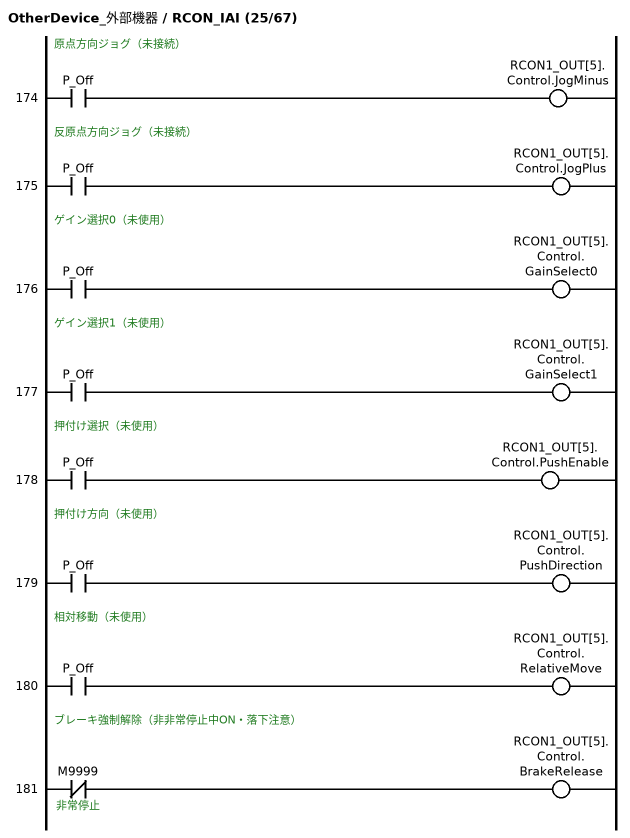
(* [picture p96: OtherDevice_外部機器 / RCON_IAI, rungs 174-181] *)
(* Rung 174: 原点方向ジョグ（未接続） *)
RCON1_OUT[5].Control.JogMinus := P_Off;
(* Rung 175: 反原点方向ジョグ（未接続） *)
RCON1_OUT[5].Control.JogPlus := P_Off;
(* Rung 176: ゲイン選択0（未使用） *)
RCON1_OUT[5].Control.GainSelect0 := P_Off;
(* Rung 177: ゲイン選択1（未使用） *)
RCON1_OUT[5].Control.GainSelect1 := P_Off;
(* Rung 178: 押付け選択（未使用） *)
RCON1_OUT[5].Control.PushEnable := P_Off;
(* Rung 179: 押付け方向（未使用） *)
RCON1_OUT[5].Control.PushDirection := P_Off;
(* Rung 180: 相対移動（未使用） *)
RCON1_OUT[5].Control.RelativeMove := P_Off;
(* Rung 181: ブレーキ強制解除（非非常停止中ON・落下注意） *)
RCON1_OUT[5].Control.BrakeRelease := NOT M9999;

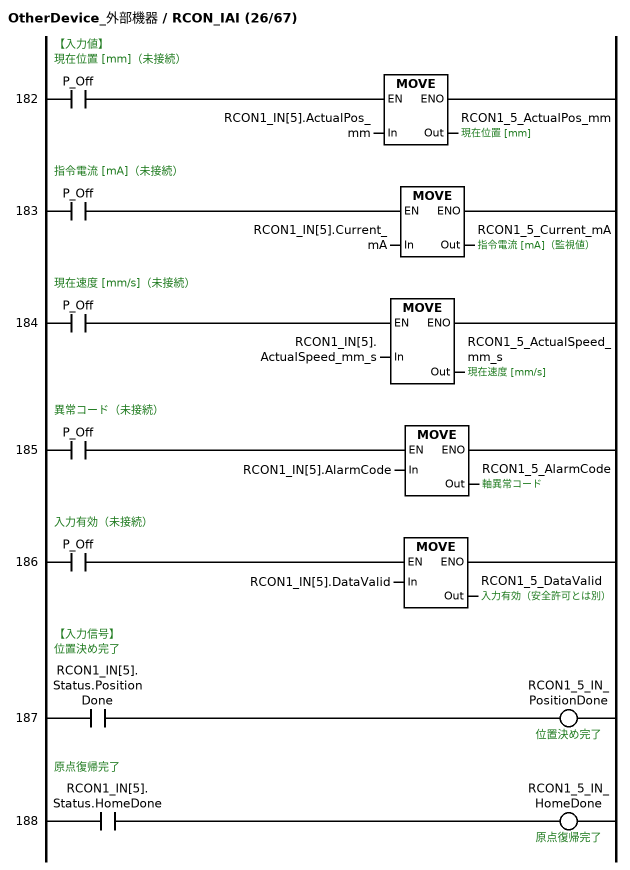
(* Rung 182: 【入力値】 / 現在位置 [mm]（未接続） *)
IF P_Off THEN RCON1_5_ActualPos_mm := RCON1_IN[5].ActualPos_mm; END_IF;
(* Rung 183: 指令電流 [mA]（未接続） *)
IF P_Off THEN RCON1_5_Current_mA := RCON1_IN[5].Current_mA; END_IF;
(* Rung 184: 現在速度 [mm/s]（未接続） *)
IF P_Off THEN RCON1_5_ActualSpeed_mm_s := RCON1_IN[5].ActualSpeed_mm_s; END_IF;
(* Rung 185: 異常コード（未接続） *)
IF P_Off THEN RCON1_5_AlarmCode := RCON1_IN[5].AlarmCode; END_IF;
(* Rung 186: 入力有効（未接続） *)
IF P_Off THEN RCON1_5_DataValid := RCON1_IN[5].DataValid; END_IF;
(* Rung 187: 【入力信号】 / 位置決め完了 *)
RCON1_5_IN_PositionDone := RCON1_IN[5].Status.PositionDone;
(* Rung 188: 原点復帰完了 *)
RCON1_5_IN_HomeDone := RCON1_IN[5].Status.HomeDone;

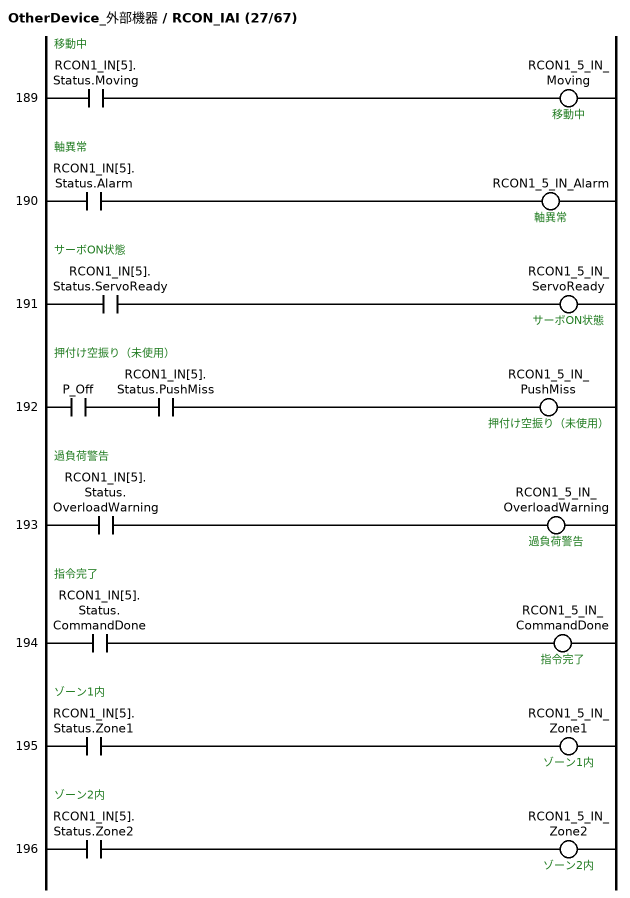
(* Rung 189: 移動中 *)
RCON1_5_IN_Moving := RCON1_IN[5].Status.Moving;
(* Rung 190: 軸異常 *)
RCON1_5_IN_Alarm := RCON1_IN[5].Status.Alarm;
(* Rung 191: サーボON状態 *)
RCON1_5_IN_ServoReady := RCON1_IN[5].Status.ServoReady;
(* Rung 192: 押付け空振り（未使用） *)
RCON1_5_IN_PushMiss := P_Off AND RCON1_IN[5].Status.PushMiss;
(* Rung 193: 過負荷警告 *)
RCON1_5_IN_OverloadWarning := RCON1_IN[5].Status.OverloadWarning;
(* Rung 194: 指令完了 *)
RCON1_5_IN_CommandDone := RCON1_IN[5].Status.CommandDone;
(* Rung 195: ゾーン1内 *)
RCON1_5_IN_Zone1 := RCON1_IN[5].Status.Zone1;
(* Rung 196: ゾーン2内 *)
RCON1_5_IN_Zone2 := RCON1_IN[5].Status.Zone2;

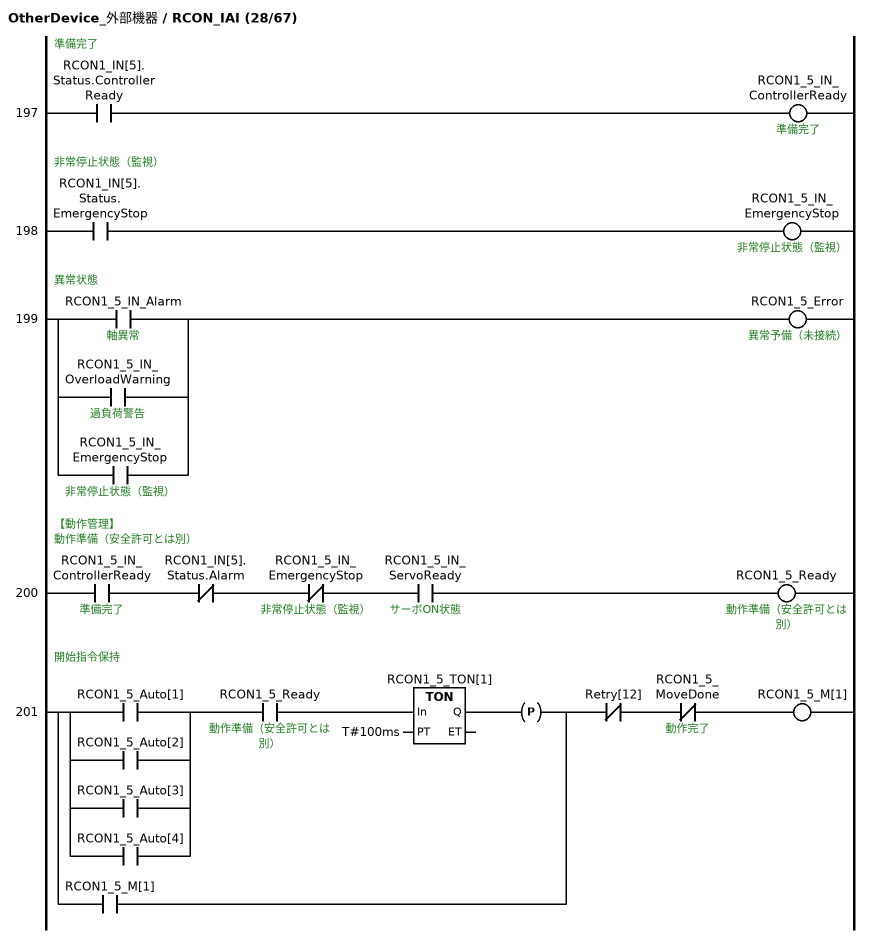
(* Rung 197: 準備完了 *)
RCON1_5_IN_ControllerReady := RCON1_IN[5].Status.ControllerReady;
(* Rung 198: 非常停止状態（監視） *)
RCON1_5_IN_EmergencyStop := RCON1_IN[5].Status.EmergencyStop;
(* Rung 199: 異常状態 *)
RCON1_5_Error := RCON1_5_IN_Alarm OR RCON1_5_IN_OverloadWarning OR RCON1_5_IN_EmergencyStop;
(* Rung 200: 【動作管理】 / 動作準備（安全許可とは別） *)
RCON1_5_Ready := RCON1_5_IN_ControllerReady AND NOT RCON1_IN[5].Status.Alarm AND NOT RCON1_5_IN_EmergencyStop AND RCON1_5_IN_ServoReady;
(* Rung 201: 開始指令保持 *)
RCON1_5_TON[1](In := (RCON1_5_Auto[1] OR RCON1_5_Auto[2] OR RCON1_5_Auto[3] OR RCON1_5_Auto[4]) AND RCON1_5_Ready, PT := T#100ms);
_e18(CLK := RCON1_5_TON[1].Q);
RCON1_5_M[1] := (_e18.Q OR RCON1_5_M[1]) AND NOT Retry[12] AND NOT RCON1_5_MoveDone;

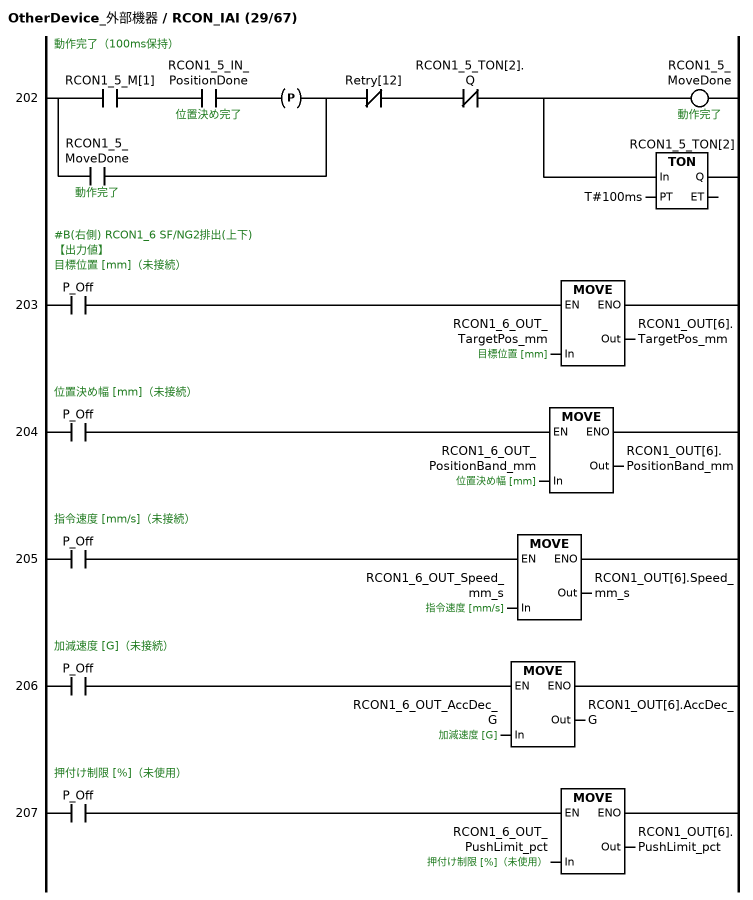
(* Rung 202: 動作完了（100ms保持） *)
_e19(CLK := RCON1_5_M[1] AND RCON1_5_IN_PositionDone);
_p20 := (_e19.Q OR RCON1_5_MoveDone) AND NOT Retry[12] AND NOT RCON1_5_TON[2].Q;
RCON1_5_MoveDone := _p20;
RCON1_5_TON[2](In := _p20, PT := T#100ms);
(* Rung 203: #B(右側) RCON1_6 SF/NG2排出(上下) / 【出力値】 / 目標位置 [mm]（未接続） *)
IF P_Off THEN RCON1_OUT[6].TargetPos_mm := RCON1_6_OUT_TargetPos_mm; END_IF;
(* Rung 204: 位置決め幅 [mm]（未接続） *)
IF P_Off THEN RCON1_OUT[6].PositionBand_mm := RCON1_6_OUT_PositionBand_mm; END_IF;
(* Rung 205: 指令速度 [mm/s]（未接続） *)
IF P_Off THEN RCON1_OUT[6].Speed_mm_s := RCON1_6_OUT_Speed_mm_s; END_IF;
(* Rung 206: 加減速度 [G]（未接続） *)
IF P_Off THEN RCON1_OUT[6].AccDec_G := RCON1_6_OUT_AccDec_G; END_IF;
(* Rung 207: 押付け制限 [%]（未使用） *)
IF P_Off THEN RCON1_OUT[6].PushLimit_pct := RCON1_6_OUT_PushLimit_pct; END_IF;

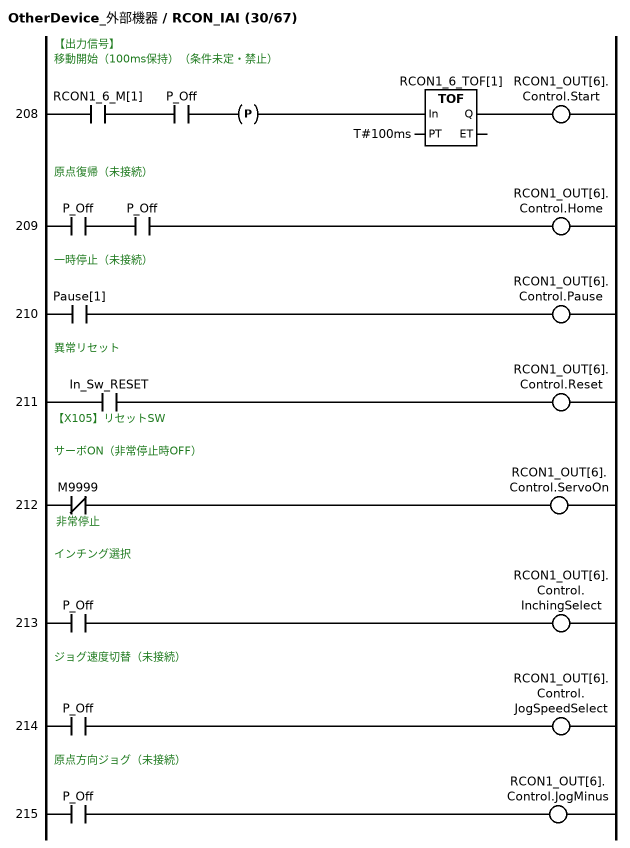
(* Rung 208: 【出力信号】 / 移動開始（100ms保持）（条件未定・禁止） *)
_e21(CLK := RCON1_6_M[1] AND P_Off);
RCON1_6_TOF[1](In := _e21.Q, PT := T#100ms);
RCON1_OUT[6].Control.Start := RCON1_6_TOF[1].Q;
(* Rung 209: 原点復帰（未接続） *)
RCON1_OUT[6].Control.Home := P_Off AND P_Off;
(* Rung 210: 一時停止（未接続） *)
RCON1_OUT[6].Control.Pause := Pause[1];
(* Rung 211: 異常リセット *)
RCON1_OUT[6].Control.Reset := In_Sw_RESET;
(* Rung 212: サーボON（非常停止時OFF） *)
RCON1_OUT[6].Control.ServoOn := NOT M9999;
(* Rung 213: インチング選択 *)
RCON1_OUT[6].Control.InchingSelect := P_Off;
(* Rung 214: ジョグ速度切替（未接続） *)
RCON1_OUT[6].Control.JogSpeedSelect := P_Off;
(* Rung 215: 原点方向ジョグ（未接続） *)
RCON1_OUT[6].Control.JogMinus := P_Off;

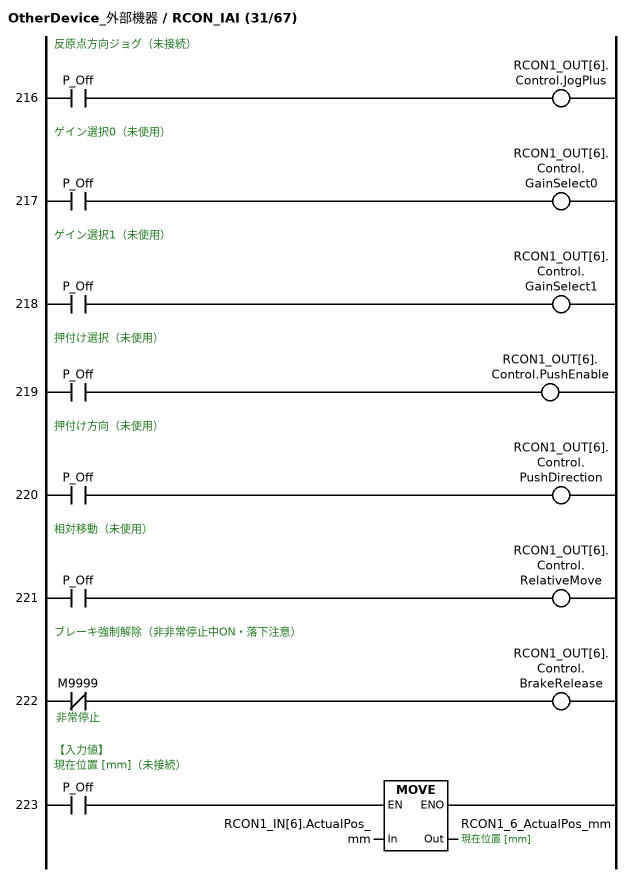
(* Rung 216: 反原点方向ジョグ（未接続） *)
RCON1_OUT[6].Control.JogPlus := P_Off;
(* Rung 217: ゲイン選択0（未使用） *)
RCON1_OUT[6].Control.GainSelect0 := P_Off;
(* Rung 218: ゲイン選択1（未使用） *)
RCON1_OUT[6].Control.GainSelect1 := P_Off;
(* Rung 219: 押付け選択（未使用） *)
RCON1_OUT[6].Control.PushEnable := P_Off;
(* Rung 220: 押付け方向（未使用） *)
RCON1_OUT[6].Control.PushDirection := P_Off;
(* Rung 221: 相対移動（未使用） *)
RCON1_OUT[6].Control.RelativeMove := P_Off;
(* Rung 222: ブレーキ強制解除（非非常停止中ON・落下注意） *)
RCON1_OUT[6].Control.BrakeRelease := NOT M9999;
(* Rung 223: 【入力値】 / 現在位置 [mm]（未接続） *)
IF P_Off THEN RCON1_6_ActualPos_mm := RCON1_IN[6].ActualPos_mm; END_IF;

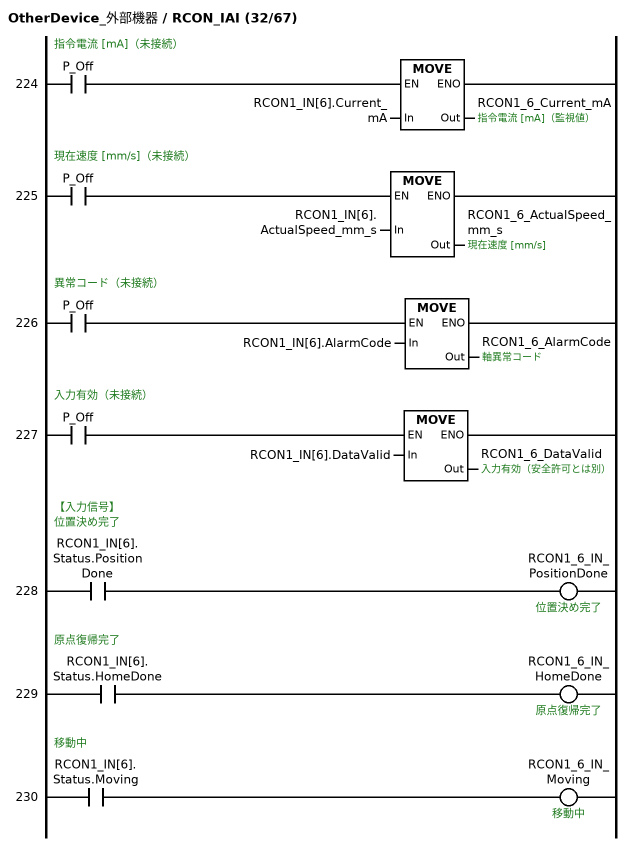
(* Rung 224: 指令電流 [mA]（未接続） *)
IF P_Off THEN RCON1_6_Current_mA := RCON1_IN[6].Current_mA; END_IF;
(* Rung 225: 現在速度 [mm/s]（未接続） *)
IF P_Off THEN RCON1_6_ActualSpeed_mm_s := RCON1_IN[6].ActualSpeed_mm_s; END_IF;
(* Rung 226: 異常コード（未接続） *)
IF P_Off THEN RCON1_6_AlarmCode := RCON1_IN[6].AlarmCode; END_IF;
(* Rung 227: 入力有効（未接続） *)
IF P_Off THEN RCON1_6_DataValid := RCON1_IN[6].DataValid; END_IF;
(* Rung 228: 【入力信号】 / 位置決め完了 *)
RCON1_6_IN_PositionDone := RCON1_IN[6].Status.PositionDone;
(* Rung 229: 原点復帰完了 *)
RCON1_6_IN_HomeDone := RCON1_IN[6].Status.HomeDone;
(* Rung 230: 移動中 *)
RCON1_6_IN_Moving := RCON1_IN[6].Status.Moving;

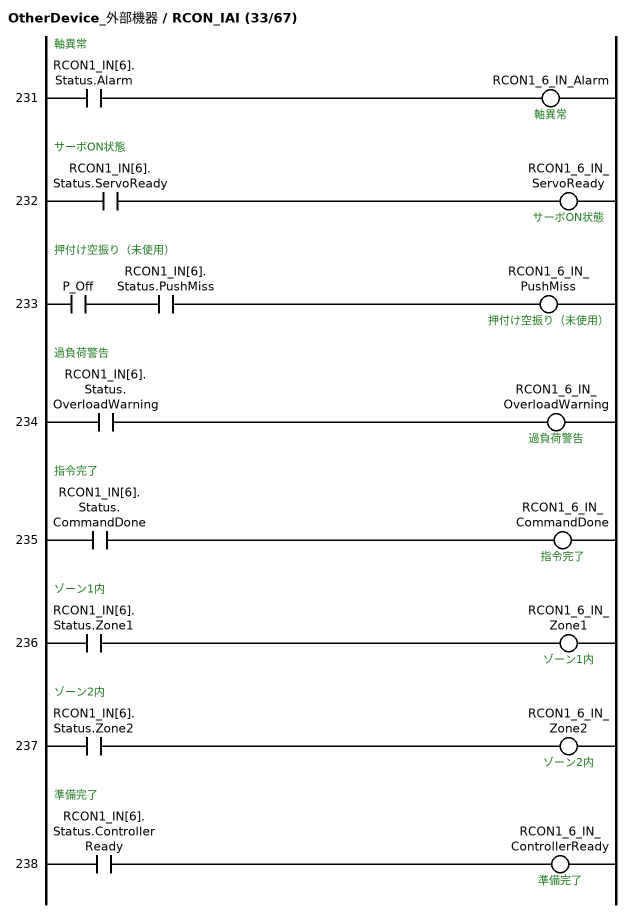
(* Rung 231: 軸異常 *)
RCON1_6_IN_Alarm := RCON1_IN[6].Status.Alarm;
(* Rung 232: サーボON状態 *)
RCON1_6_IN_ServoReady := RCON1_IN[6].Status.ServoReady;
(* Rung 233: 押付け空振り（未使用） *)
RCON1_6_IN_PushMiss := P_Off AND RCON1_IN[6].Status.PushMiss;
(* Rung 234: 過負荷警告 *)
RCON1_6_IN_OverloadWarning := RCON1_IN[6].Status.OverloadWarning;
(* Rung 235: 指令完了 *)
RCON1_6_IN_CommandDone := RCON1_IN[6].Status.CommandDone;
(* Rung 236: ゾーン1内 *)
RCON1_6_IN_Zone1 := RCON1_IN[6].Status.Zone1;
(* Rung 237: ゾーン2内 *)
RCON1_6_IN_Zone2 := RCON1_IN[6].Status.Zone2;
(* Rung 238: 準備完了 *)
RCON1_6_IN_ControllerReady := RCON1_IN[6].Status.ControllerReady;

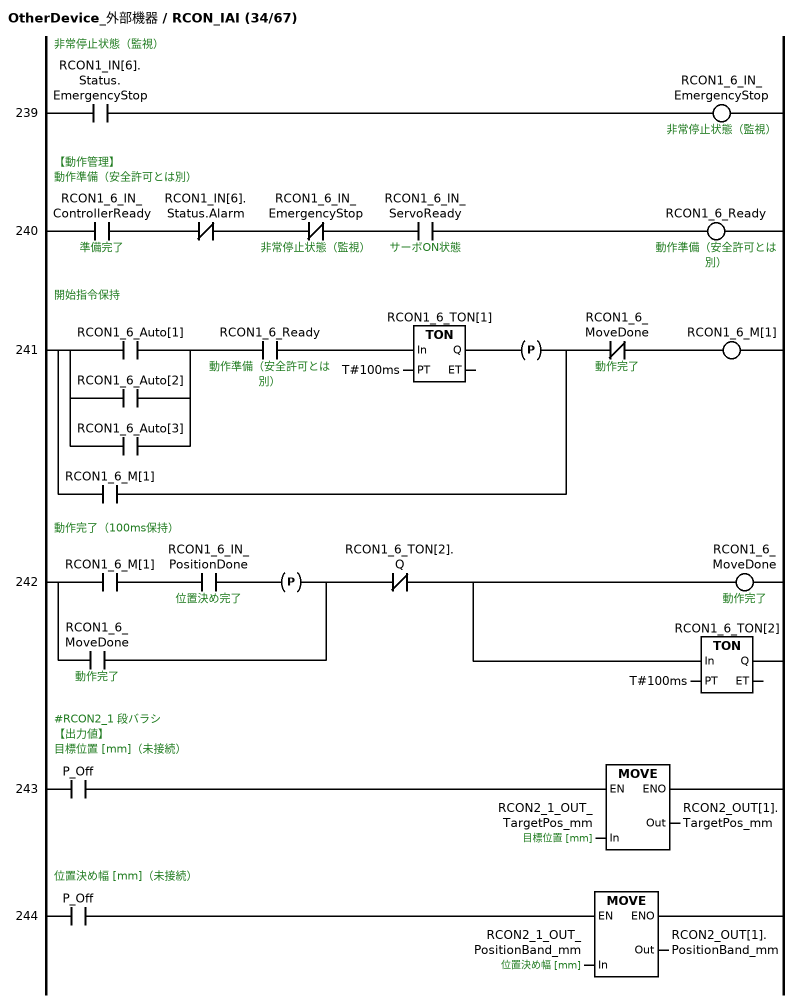
(* Rung 239: 非常停止状態（監視） *)
RCON1_6_IN_EmergencyStop := RCON1_IN[6].Status.EmergencyStop;
(* Rung 240: 【動作管理】 / 動作準備（安全許可とは別） *)
RCON1_6_Ready := RCON1_6_IN_ControllerReady AND NOT RCON1_IN[6].Status.Alarm AND NOT RCON1_6_IN_EmergencyStop AND RCON1_6_IN_ServoReady;
(* Rung 241: 開始指令保持 *)
RCON1_6_TON[1](In := (RCON1_6_Auto[1] OR RCON1_6_Auto[2] OR RCON1_6_Auto[3]) AND RCON1_6_Ready, PT := T#100ms);
_e22(CLK := RCON1_6_TON[1].Q);
RCON1_6_M[1] := (_e22.Q OR RCON1_6_M[1]) AND NOT RCON1_6_MoveDone;
(* Rung 242: 動作完了（100ms保持） *)
_e23(CLK := RCON1_6_M[1] AND RCON1_6_IN_PositionDone);
_p24 := (_e23.Q OR RCON1_6_MoveDone) AND NOT RCON1_6_TON[2].Q;
RCON1_6_MoveDone := _p24;
RCON1_6_TON[2](In := _p24, PT := T#100ms);
(* Rung 243: #RCON2_1 段バラシ / 【出力値】 / 目標位置 [mm]（未接続） *)
IF P_Off THEN RCON2_OUT[1].TargetPos_mm := RCON2_1_OUT_TargetPos_mm; END_IF;
(* Rung 244: 位置決め幅 [mm]（未接続） *)
IF P_Off THEN RCON2_OUT[1].PositionBand_mm := RCON2_1_OUT_PositionBand_mm; END_IF;

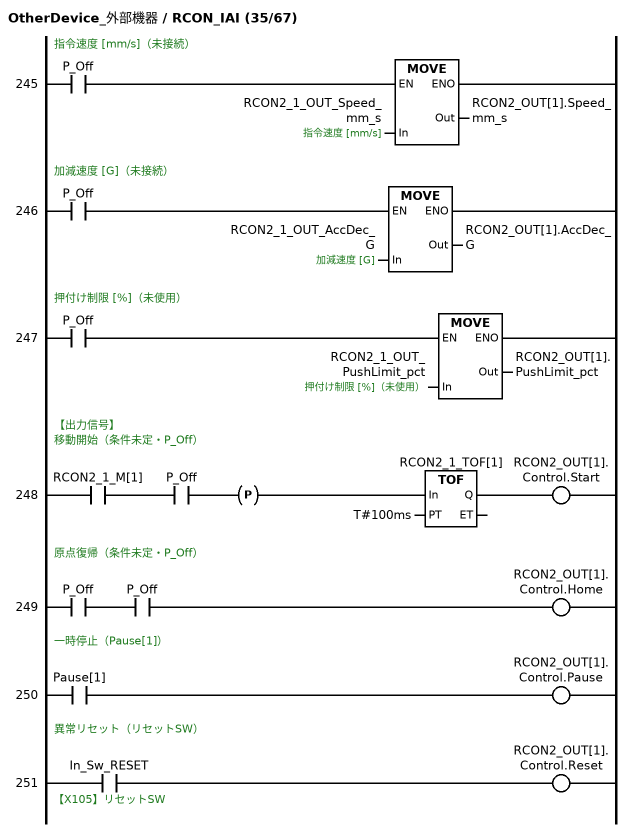
(* Rung 245: 指令速度 [mm/s]（未接続） *)
IF P_Off THEN RCON2_OUT[1].Speed_mm_s := RCON2_1_OUT_Speed_mm_s; END_IF;
(* Rung 246: 加減速度 [G]（未接続） *)
IF P_Off THEN RCON2_OUT[1].AccDec_G := RCON2_1_OUT_AccDec_G; END_IF;
(* Rung 247: 押付け制限 [%]（未使用） *)
IF P_Off THEN RCON2_OUT[1].PushLimit_pct := RCON2_1_OUT_PushLimit_pct; END_IF;
(* Rung 248: 【出力信号】 / 移動開始（条件未定・P_Off） *)
_e25(CLK := RCON2_1_M[1] AND P_Off);
RCON2_1_TOF[1](In := _e25.Q, PT := T#100ms);
RCON2_OUT[1].Control.Start := RCON2_1_TOF[1].Q;
(* Rung 249: 原点復帰（条件未定・P_Off） *)
RCON2_OUT[1].Control.Home := P_Off AND P_Off;
(* Rung 250: 一時停止（Pause[1]） *)
RCON2_OUT[1].Control.Pause := Pause[1];
(* Rung 251: 異常リセット（リセットSW） *)
RCON2_OUT[1].Control.Reset := In_Sw_RESET;

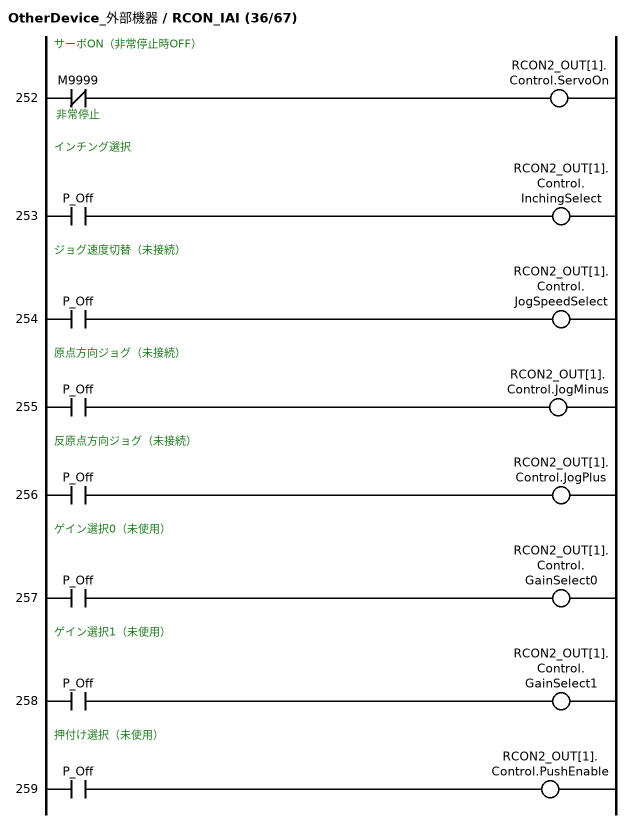
(* Rung 252: サーボON（非常停止時OFF） *)
RCON2_OUT[1].Control.ServoOn := NOT M9999;
(* Rung 253: インチング選択 *)
RCON2_OUT[1].Control.InchingSelect := P_Off;
(* Rung 254: ジョグ速度切替（未接続） *)
RCON2_OUT[1].Control.JogSpeedSelect := P_Off;
(* Rung 255: 原点方向ジョグ（未接続） *)
RCON2_OUT[1].Control.JogMinus := P_Off;
(* Rung 256: 反原点方向ジョグ（未接続） *)
RCON2_OUT[1].Control.JogPlus := P_Off;
(* Rung 257: ゲイン選択0（未使用） *)
RCON2_OUT[1].Control.GainSelect0 := P_Off;
(* Rung 258: ゲイン選択1（未使用） *)
RCON2_OUT[1].Control.GainSelect1 := P_Off;
(* Rung 259: 押付け選択（未使用） *)
RCON2_OUT[1].Control.PushEnable := P_Off;

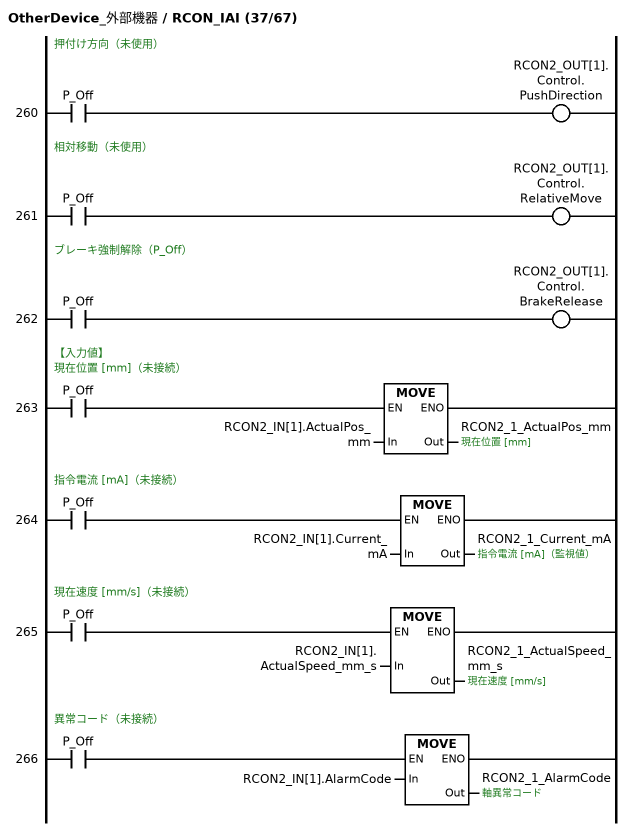
(* Rung 260: 押付け方向（未使用） *)
RCON2_OUT[1].Control.PushDirection := P_Off;
(* Rung 261: 相対移動（未使用） *)
RCON2_OUT[1].Control.RelativeMove := P_Off;
(* Rung 262: ブレーキ強制解除（P_Off） *)
RCON2_OUT[1].Control.BrakeRelease := P_Off;
(* Rung 263: 【入力値】 / 現在位置 [mm]（未接続） *)
IF P_Off THEN RCON2_1_ActualPos_mm := RCON2_IN[1].ActualPos_mm; END_IF;
(* Rung 264: 指令電流 [mA]（未接続） *)
IF P_Off THEN RCON2_1_Current_mA := RCON2_IN[1].Current_mA; END_IF;
(* Rung 265: 現在速度 [mm/s]（未接続） *)
IF P_Off THEN RCON2_1_ActualSpeed_mm_s := RCON2_IN[1].ActualSpeed_mm_s; END_IF;
(* Rung 266: 異常コード（未接続） *)
IF P_Off THEN RCON2_1_AlarmCode := RCON2_IN[1].AlarmCode; END_IF;

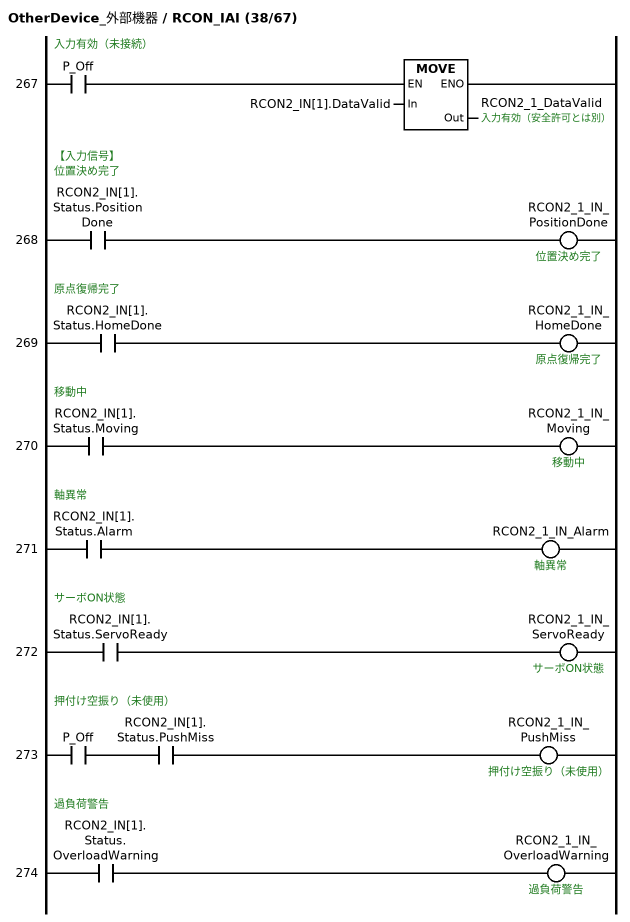
(* Rung 267: 入力有効（未接続） *)
IF P_Off THEN RCON2_1_DataValid := RCON2_IN[1].DataValid; END_IF;
(* Rung 268: 【入力信号】 / 位置決め完了 *)
RCON2_1_IN_PositionDone := RCON2_IN[1].Status.PositionDone;
(* Rung 269: 原点復帰完了 *)
RCON2_1_IN_HomeDone := RCON2_IN[1].Status.HomeDone;
(* Rung 270: 移動中 *)
RCON2_1_IN_Moving := RCON2_IN[1].Status.Moving;
(* Rung 271: 軸異常 *)
RCON2_1_IN_Alarm := RCON2_IN[1].Status.Alarm;
(* Rung 272: サーボON状態 *)
RCON2_1_IN_ServoReady := RCON2_IN[1].Status.ServoReady;
(* Rung 273: 押付け空振り（未使用） *)
RCON2_1_IN_PushMiss := P_Off AND RCON2_IN[1].Status.PushMiss;
(* Rung 274: 過負荷警告 *)
RCON2_1_IN_OverloadWarning := RCON2_IN[1].Status.OverloadWarning;

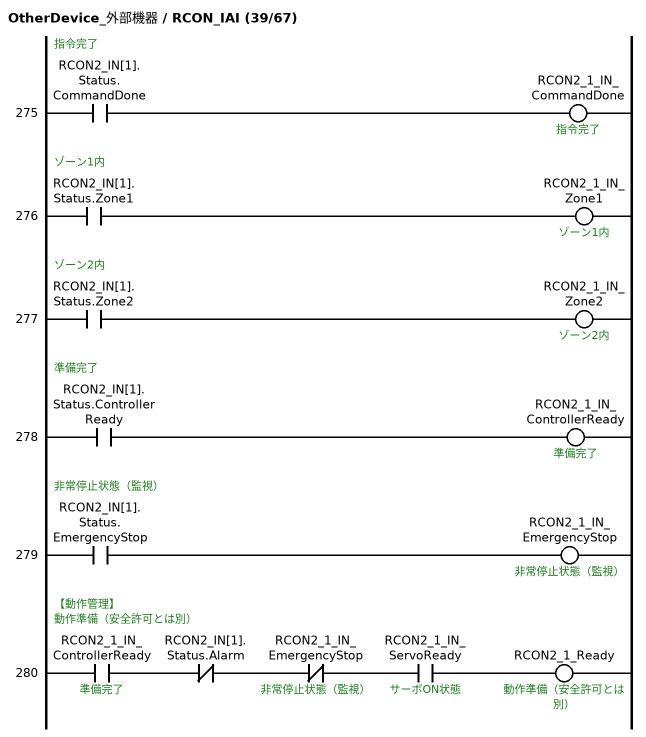
(* Rung 275: 指令完了 *)
RCON2_1_IN_CommandDone := RCON2_IN[1].Status.CommandDone;
(* Rung 276: ゾーン1内 *)
RCON2_1_IN_Zone1 := RCON2_IN[1].Status.Zone1;
(* Rung 277: ゾーン2内 *)
RCON2_1_IN_Zone2 := RCON2_IN[1].Status.Zone2;
(* Rung 278: 準備完了 *)
RCON2_1_IN_ControllerReady := RCON2_IN[1].Status.ControllerReady;
(* Rung 279: 非常停止状態（監視） *)
RCON2_1_IN_EmergencyStop := RCON2_IN[1].Status.EmergencyStop;
(* Rung 280: 【動作管理】 / 動作準備（安全許可とは別） *)
RCON2_1_Ready := RCON2_1_IN_ControllerReady AND NOT RCON2_IN[1].Status.Alarm AND NOT RCON2_1_IN_EmergencyStop AND RCON2_1_IN_ServoReady;

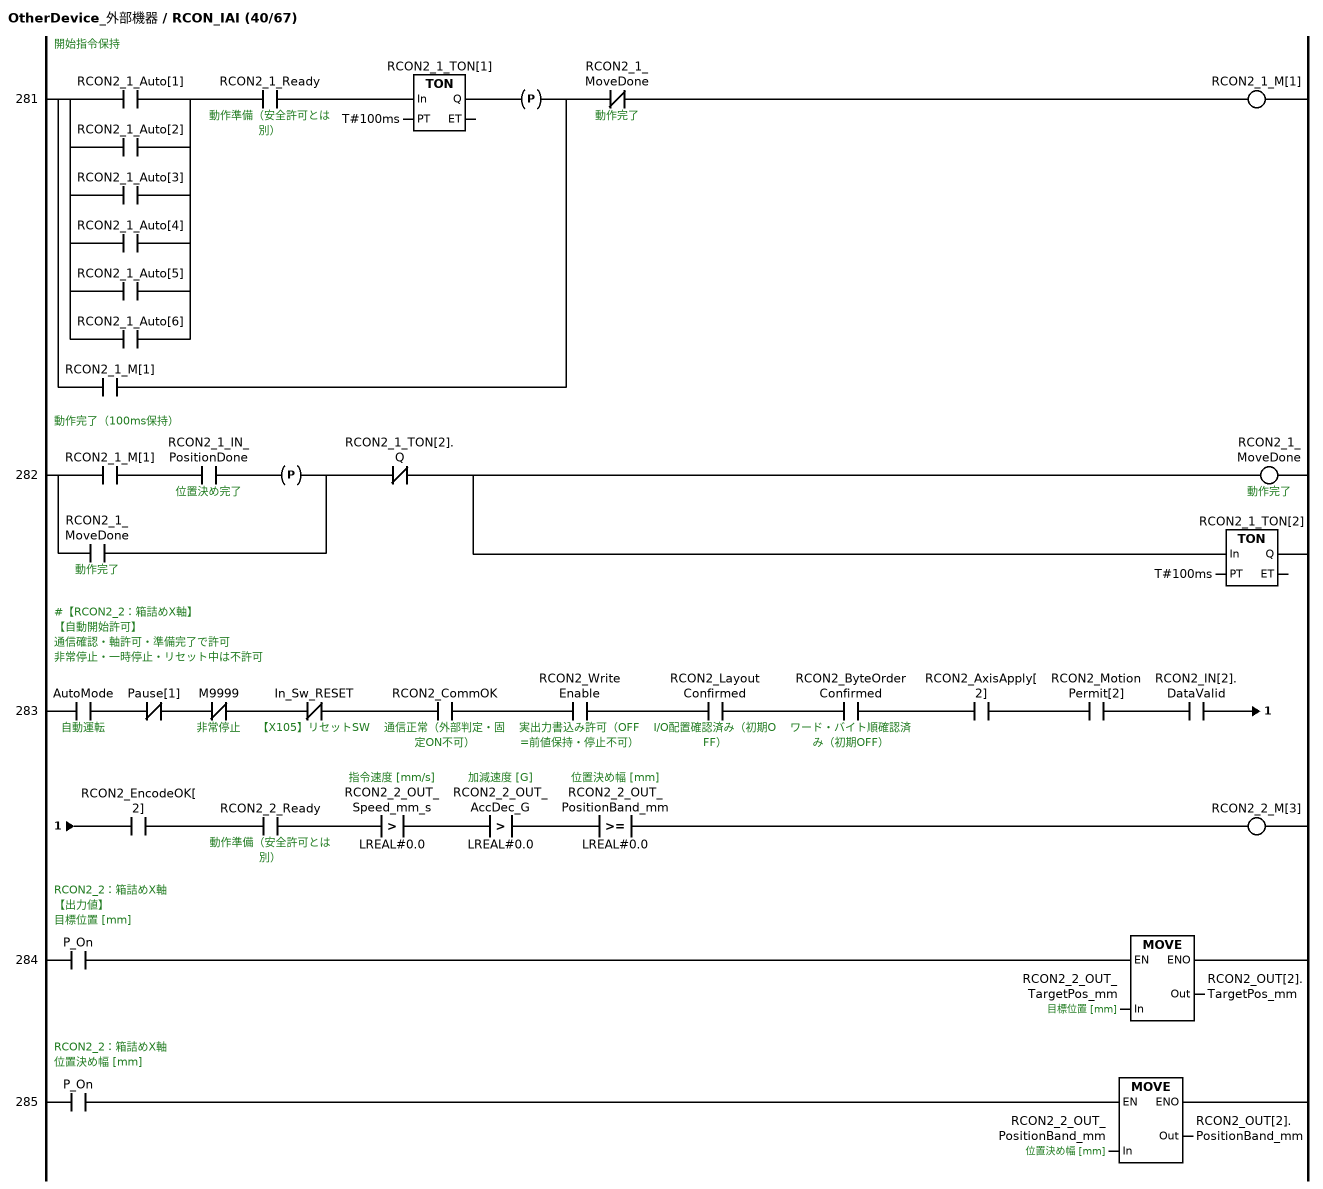
(* Rung 281: 開始指令保持 *)
RCON2_1_TON[1](In := (RCON2_1_Auto[1] OR RCON2_1_Auto[2] OR RCON2_1_Auto[3] OR RCON2_1_Auto[4] OR RCON2_1_Auto[5] OR RCON2_1_Auto[6]) AND RCON2_1_Ready, PT := T#100ms);
_e26(CLK := RCON2_1_TON[1].Q);
RCON2_1_M[1] := (_e26.Q OR RCON2_1_M[1]) AND NOT RCON2_1_MoveDone;
(* Rung 282: 動作完了（100ms保持） *)
_e27(CLK := RCON2_1_M[1] AND RCON2_1_IN_PositionDone);
_p28 := (_e27.Q OR RCON2_1_MoveDone) AND NOT RCON2_1_TON[2].Q;
RCON2_1_MoveDone := _p28;
RCON2_1_TON[2](In := _p28, PT := T#100ms);
(* Rung 283: #【RCON2_2：箱詰めX軸】 / 【自動開始許可】 / 通信確認・軸許可・準備完了で許可 / 非常停止・一時停止・リセット中は不許可 *)
RCON2_2_M[3] := AutoMode AND NOT Pause[1] AND NOT M9999 AND NOT In_Sw_RESET AND RCON2_CommOK AND RCON2_WriteEnable AND RCON2_LayoutConfirmed AND RCON2_ByteOrderConfirmed AND RCON2_AxisApply[2] AND RCON2_MotionPermit[2] AND RCON2_IN[2].DataValid AND RCON2_EncodeOK[2] AND RCON2_2_Ready AND (RCON2_2_OUT_Speed_mm_s > LREAL#0.0) AND (RCON2_2_OUT_AccDec_G > LREAL#0.0) AND (RCON2_2_OUT_PositionBand_mm >= LREAL#0.0);
(* Rung 284: RCON2_2：箱詰めX軸 / 【出力値】 / 目標位置 [mm] *)
IF P_On THEN RCON2_OUT[2].TargetPos_mm := RCON2_2_OUT_TargetPos_mm; END_IF;
(* Rung 285: RCON2_2：箱詰めX軸 / 位置決め幅 [mm] *)
IF P_On THEN RCON2_OUT[2].PositionBand_mm := RCON2_2_OUT_PositionBand_mm; END_IF;

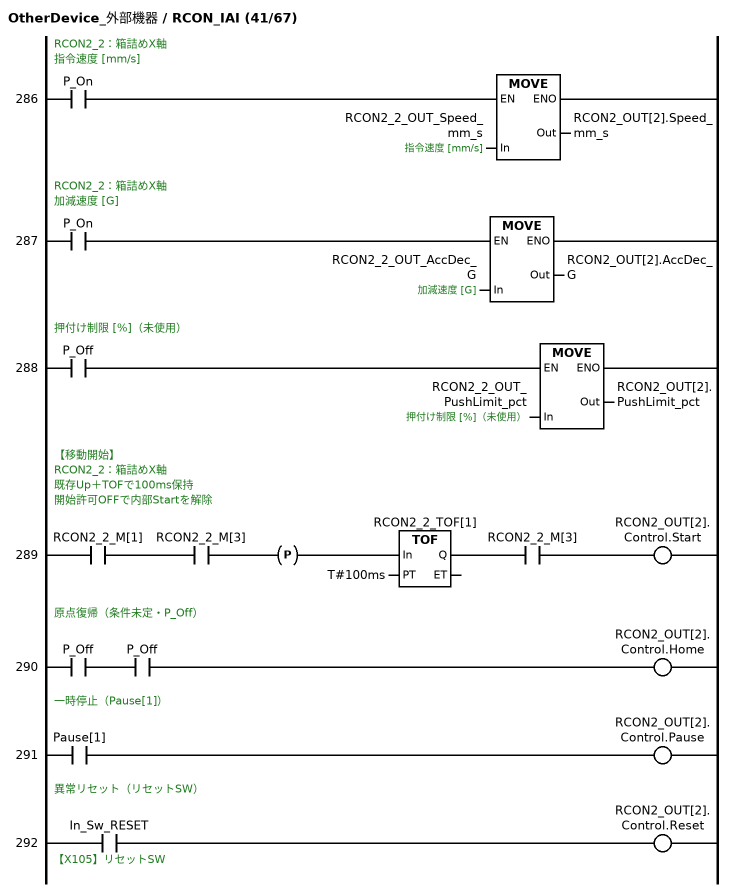
(* Rung 286: RCON2_2：箱詰めX軸 / 指令速度 [mm/s] *)
IF P_On THEN RCON2_OUT[2].Speed_mm_s := RCON2_2_OUT_Speed_mm_s; END_IF;
(* Rung 287: RCON2_2：箱詰めX軸 / 加減速度 [G] *)
IF P_On THEN RCON2_OUT[2].AccDec_G := RCON2_2_OUT_AccDec_G; END_IF;
(* Rung 288: 押付け制限 [%]（未使用） *)
IF P_Off THEN RCON2_OUT[2].PushLimit_pct := RCON2_2_OUT_PushLimit_pct; END_IF;
(* Rung 289: 【移動開始】 / RCON2_2：箱詰めX軸 / 既存Up＋TOFで100ms保持 / 開始許可OFFで内部Startを解除 *)
_e29(CLK := RCON2_2_M[1] AND RCON2_2_M[3]);
RCON2_2_TOF[1](In := _e29.Q, PT := T#100ms);
RCON2_OUT[2].Control.Start := RCON2_2_TOF[1].Q AND RCON2_2_M[3];
(* Rung 290: 原点復帰（条件未定・P_Off） *)
RCON2_OUT[2].Control.Home := P_Off AND P_Off;
(* Rung 291: 一時停止（Pause[1]） *)
RCON2_OUT[2].Control.Pause := Pause[1];
(* Rung 292: 異常リセット（リセットSW） *)
RCON2_OUT[2].Control.Reset := In_Sw_RESET;

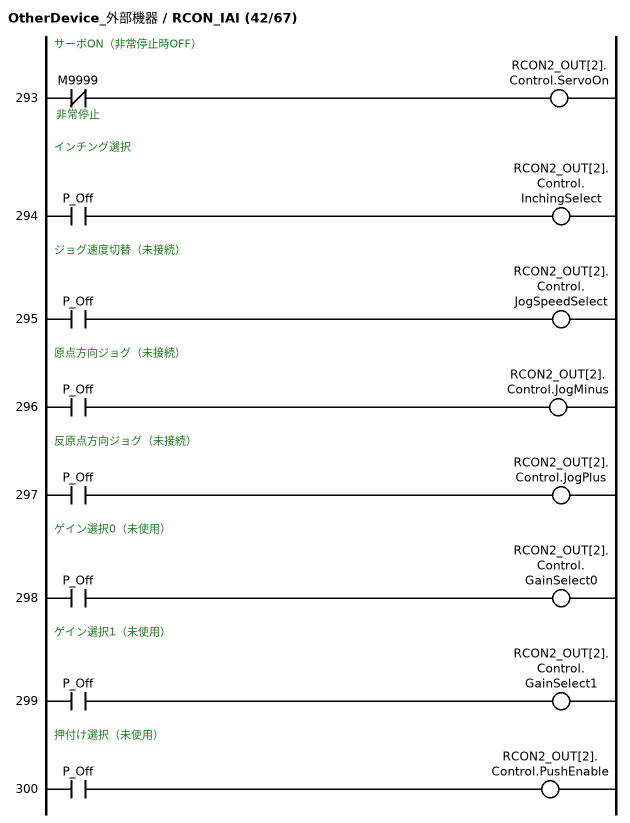
(* Rung 293: サーボON（非常停止時OFF） *)
RCON2_OUT[2].Control.ServoOn := NOT M9999;
(* Rung 294: インチング選択 *)
RCON2_OUT[2].Control.InchingSelect := P_Off;
(* Rung 295: ジョグ速度切替（未接続） *)
RCON2_OUT[2].Control.JogSpeedSelect := P_Off;
(* Rung 296: 原点方向ジョグ（未接続） *)
RCON2_OUT[2].Control.JogMinus := P_Off;
(* Rung 297: 反原点方向ジョグ（未接続） *)
RCON2_OUT[2].Control.JogPlus := P_Off;
(* Rung 298: ゲイン選択0（未使用） *)
RCON2_OUT[2].Control.GainSelect0 := P_Off;
(* Rung 299: ゲイン選択1（未使用） *)
RCON2_OUT[2].Control.GainSelect1 := P_Off;
(* Rung 300: 押付け選択（未使用） *)
RCON2_OUT[2].Control.PushEnable := P_Off;

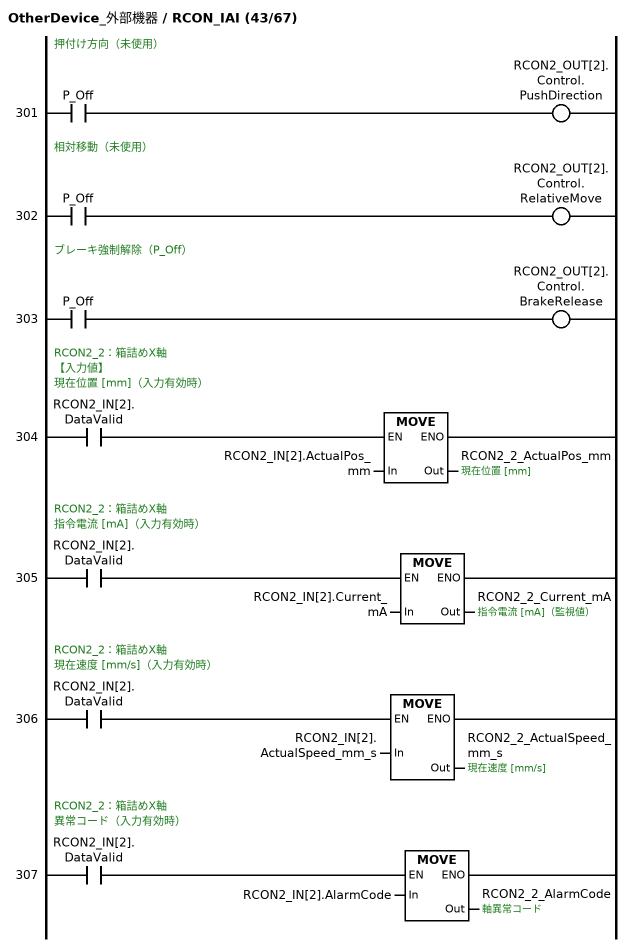
(* Rung 301: 押付け方向（未使用） *)
RCON2_OUT[2].Control.PushDirection := P_Off;
(* Rung 302: 相対移動（未使用） *)
RCON2_OUT[2].Control.RelativeMove := P_Off;
(* Rung 303: ブレーキ強制解除（P_Off） *)
RCON2_OUT[2].Control.BrakeRelease := P_Off;
(* Rung 304: RCON2_2：箱詰めX軸 / 【入力値】 / 現在位置 [mm]（入力有効時） *)
IF RCON2_IN[2].DataValid THEN RCON2_2_ActualPos_mm := RCON2_IN[2].ActualPos_mm; END_IF;
(* Rung 305: RCON2_2：箱詰めX軸 / 指令電流 [mA]（入力有効時） *)
IF RCON2_IN[2].DataValid THEN RCON2_2_Current_mA := RCON2_IN[2].Current_mA; END_IF;
(* Rung 306: RCON2_2：箱詰めX軸 / 現在速度 [mm/s]（入力有効時） *)
IF RCON2_IN[2].DataValid THEN RCON2_2_ActualSpeed_mm_s := RCON2_IN[2].ActualSpeed_mm_s; END_IF;
(* Rung 307: RCON2_2：箱詰めX軸 / 異常コード（入力有効時） *)
IF RCON2_IN[2].DataValid THEN RCON2_2_AlarmCode := RCON2_IN[2].AlarmCode; END_IF;

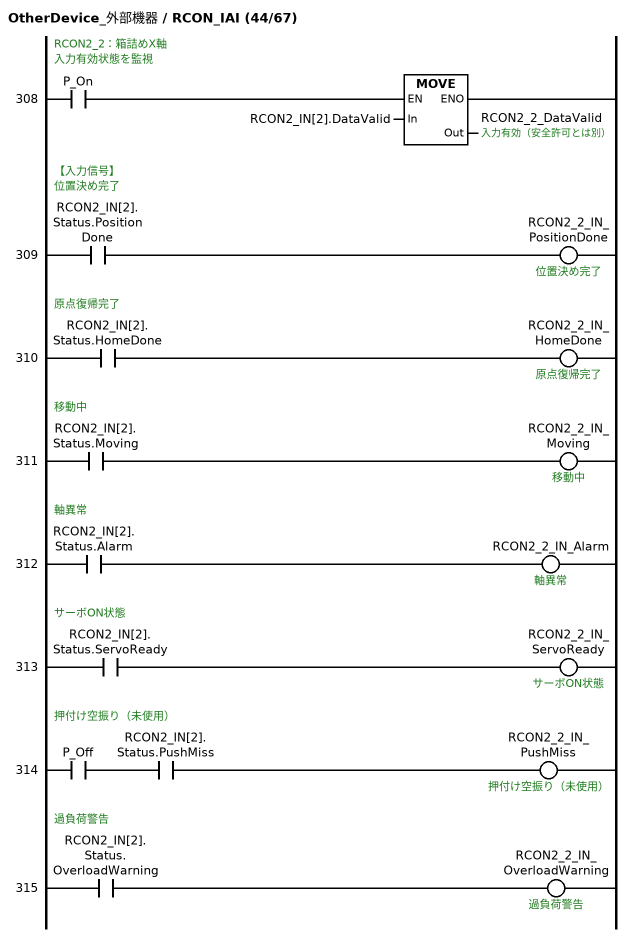
(* Rung 308: RCON2_2：箱詰めX軸 / 入力有効状態を監視 *)
IF P_On THEN RCON2_2_DataValid := RCON2_IN[2].DataValid; END_IF;
(* Rung 309: 【入力信号】 / 位置決め完了 *)
RCON2_2_IN_PositionDone := RCON2_IN[2].Status.PositionDone;
(* Rung 310: 原点復帰完了 *)
RCON2_2_IN_HomeDone := RCON2_IN[2].Status.HomeDone;
(* Rung 311: 移動中 *)
RCON2_2_IN_Moving := RCON2_IN[2].Status.Moving;
(* Rung 312: 軸異常 *)
RCON2_2_IN_Alarm := RCON2_IN[2].Status.Alarm;
(* Rung 313: サーボON状態 *)
RCON2_2_IN_ServoReady := RCON2_IN[2].Status.ServoReady;
(* Rung 314: 押付け空振り（未使用） *)
RCON2_2_IN_PushMiss := P_Off AND RCON2_IN[2].Status.PushMiss;
(* Rung 315: 過負荷警告 *)
RCON2_2_IN_OverloadWarning := RCON2_IN[2].Status.OverloadWarning;

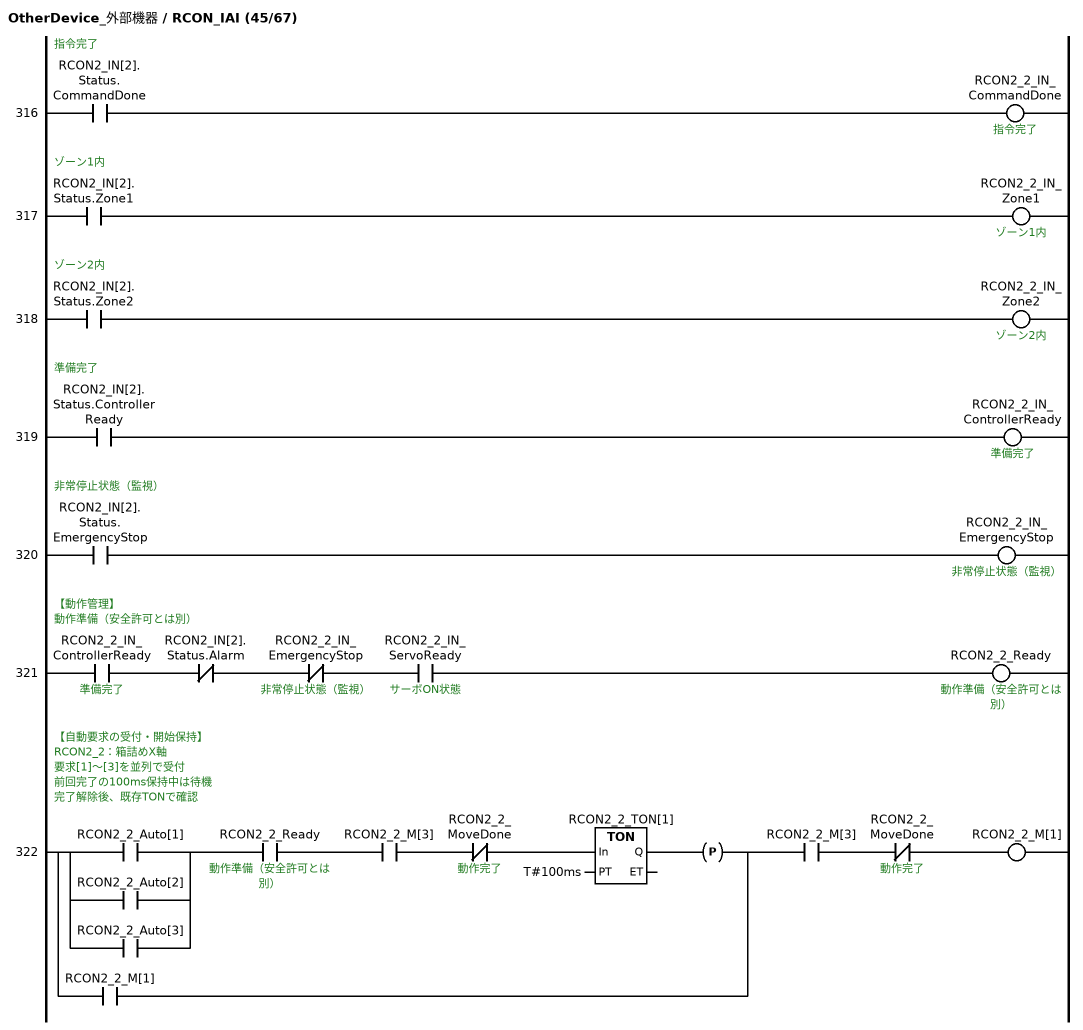
(* Rung 316: 指令完了 *)
RCON2_2_IN_CommandDone := RCON2_IN[2].Status.CommandDone;
(* Rung 317: ゾーン1内 *)
RCON2_2_IN_Zone1 := RCON2_IN[2].Status.Zone1;
(* Rung 318: ゾーン2内 *)
RCON2_2_IN_Zone2 := RCON2_IN[2].Status.Zone2;
(* Rung 319: 準備完了 *)
RCON2_2_IN_ControllerReady := RCON2_IN[2].Status.ControllerReady;
(* Rung 320: 非常停止状態（監視） *)
RCON2_2_IN_EmergencyStop := RCON2_IN[2].Status.EmergencyStop;
(* Rung 321: 【動作管理】 / 動作準備（安全許可とは別） *)
RCON2_2_Ready := RCON2_2_IN_ControllerReady AND NOT RCON2_IN[2].Status.Alarm AND NOT RCON2_2_IN_EmergencyStop AND RCON2_2_IN_ServoReady;
(* Rung 322: 【自動要求の受付・開始保持】 / RCON2_2：箱詰めX軸 / 要求[1]～[3]を並列で受付 / 前回完了の100ms保持中は待機 / 完了解除後、既存TONで確認 *)
RCON2_2_TON[1](In := (RCON2_2_Auto[1] OR RCON2_2_Auto[2] OR RCON2_2_Auto[3]) AND RCON2_2_Ready AND RCON2_2_M[3] AND NOT RCON2_2_MoveDone, PT := T#100ms);
_e30(CLK := RCON2_2_TON[1].Q);
RCON2_2_M[1] := (_e30.Q OR RCON2_2_M[1]) AND RCON2_2_M[3] AND NOT RCON2_2_MoveDone;

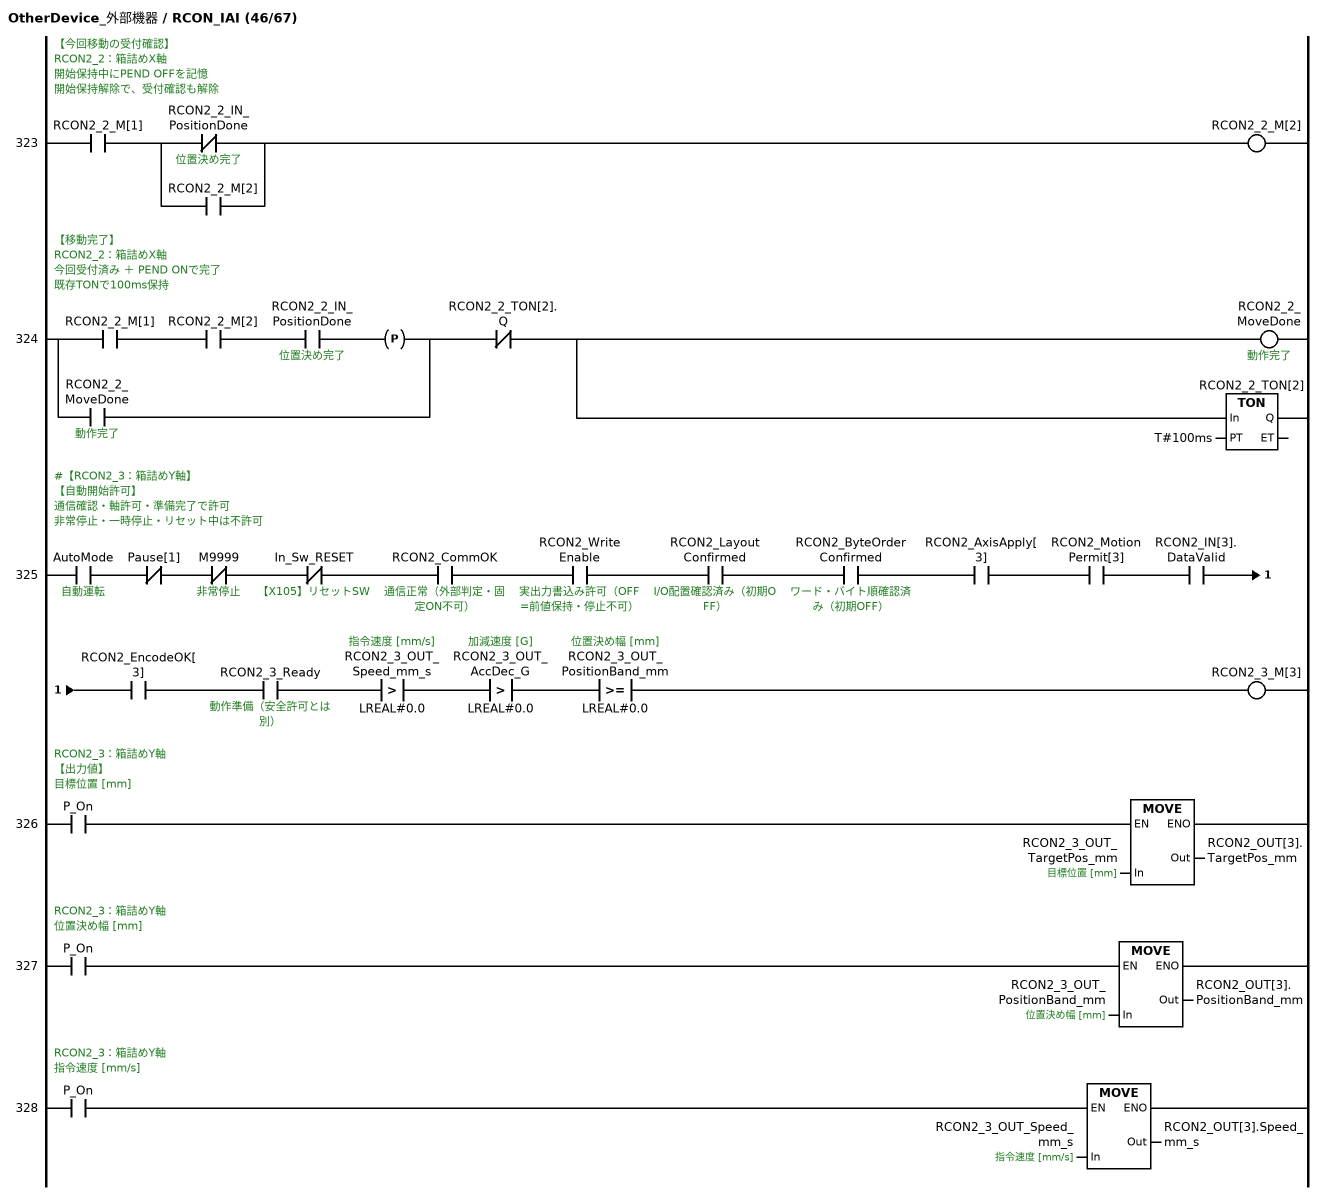
(* Rung 323: 【今回移動の受付確認】 / RCON2_2：箱詰めX軸 / 開始保持中にPEND OFFを記憶 / 開始保持解除で、受付確認も解除 *)
RCON2_2_M[2] := RCON2_2_M[1] AND (NOT RCON2_2_IN_PositionDone OR RCON2_2_M[2]);
(* Rung 324: 【移動完了】 / RCON2_2：箱詰めX軸 / 今回受付済み ＋ PEND ONで完了 / 既存TONで100ms保持 *)
_e31(CLK := RCON2_2_M[1] AND RCON2_2_M[2] AND RCON2_2_IN_PositionDone);
_p32 := (_e31.Q OR RCON2_2_MoveDone) AND NOT RCON2_2_TON[2].Q;
RCON2_2_MoveDone := _p32;
RCON2_2_TON[2](In := _p32, PT := T#100ms);
(* Rung 325: #【RCON2_3：箱詰めY軸】 / 【自動開始許可】 / 通信確認・軸許可・準備完了で許可 / 非常停止・一時停止・リセット中は不許可 *)
RCON2_3_M[3] := AutoMode AND NOT Pause[1] AND NOT M9999 AND NOT In_Sw_RESET AND RCON2_CommOK AND RCON2_WriteEnable AND RCON2_LayoutConfirmed AND RCON2_ByteOrderConfirmed AND RCON2_AxisApply[3] AND RCON2_MotionPermit[3] AND RCON2_IN[3].DataValid AND RCON2_EncodeOK[3] AND RCON2_3_Ready AND (RCON2_3_OUT_Speed_mm_s > LREAL#0.0) AND (RCON2_3_OUT_AccDec_G > LREAL#0.0) AND (RCON2_3_OUT_PositionBand_mm >= LREAL#0.0);
(* Rung 326: RCON2_3：箱詰めY軸 / 【出力値】 / 目標位置 [mm] *)
IF P_On THEN RCON2_OUT[3].TargetPos_mm := RCON2_3_OUT_TargetPos_mm; END_IF;
(* Rung 327: RCON2_3：箱詰めY軸 / 位置決め幅 [mm] *)
IF P_On THEN RCON2_OUT[3].PositionBand_mm := RCON2_3_OUT_PositionBand_mm; END_IF;
(* Rung 328: RCON2_3：箱詰めY軸 / 指令速度 [mm/s] *)
IF P_On THEN RCON2_OUT[3].Speed_mm_s := RCON2_3_OUT_Speed_mm_s; END_IF;

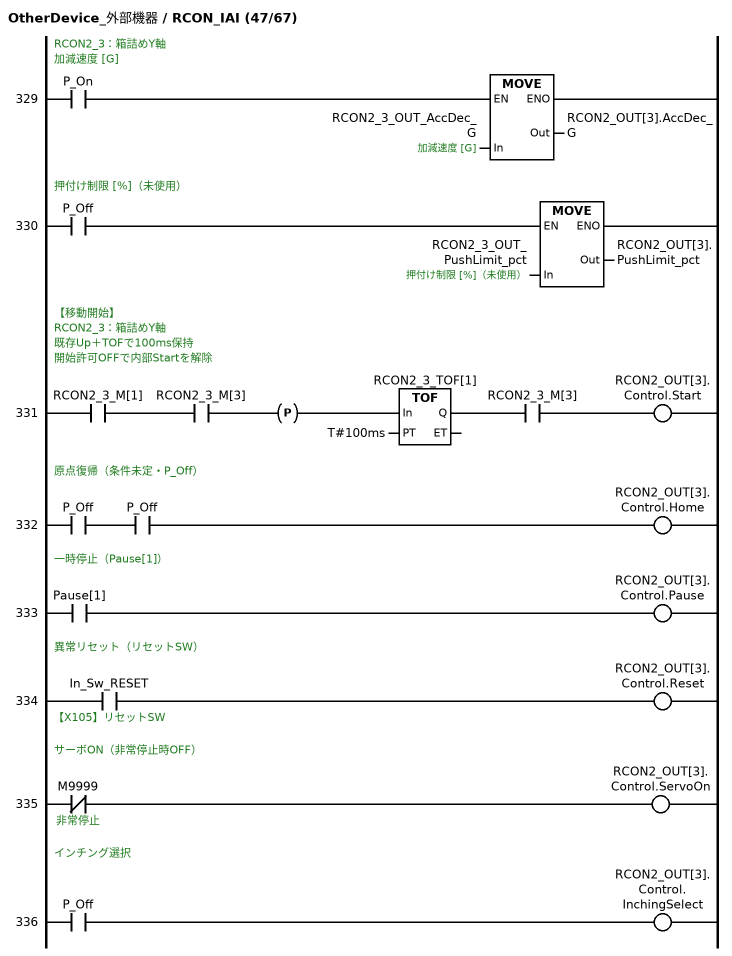
(* Rung 329: RCON2_3：箱詰めY軸 / 加減速度 [G] *)
IF P_On THEN RCON2_OUT[3].AccDec_G := RCON2_3_OUT_AccDec_G; END_IF;
(* Rung 330: 押付け制限 [%]（未使用） *)
IF P_Off THEN RCON2_OUT[3].PushLimit_pct := RCON2_3_OUT_PushLimit_pct; END_IF;
(* Rung 331: 【移動開始】 / RCON2_3：箱詰めY軸 / 既存Up＋TOFで100ms保持 / 開始許可OFFで内部Startを解除 *)
_e33(CLK := RCON2_3_M[1] AND RCON2_3_M[3]);
RCON2_3_TOF[1](In := _e33.Q, PT := T#100ms);
RCON2_OUT[3].Control.Start := RCON2_3_TOF[1].Q AND RCON2_3_M[3];
(* Rung 332: 原点復帰（条件未定・P_Off） *)
RCON2_OUT[3].Control.Home := P_Off AND P_Off;
(* Rung 333: 一時停止（Pause[1]） *)
RCON2_OUT[3].Control.Pause := Pause[1];
(* Rung 334: 異常リセット（リセットSW） *)
RCON2_OUT[3].Control.Reset := In_Sw_RESET;
(* Rung 335: サーボON（非常停止時OFF） *)
RCON2_OUT[3].Control.ServoOn := NOT M9999;
(* Rung 336: インチング選択 *)
RCON2_OUT[3].Control.InchingSelect := P_Off;

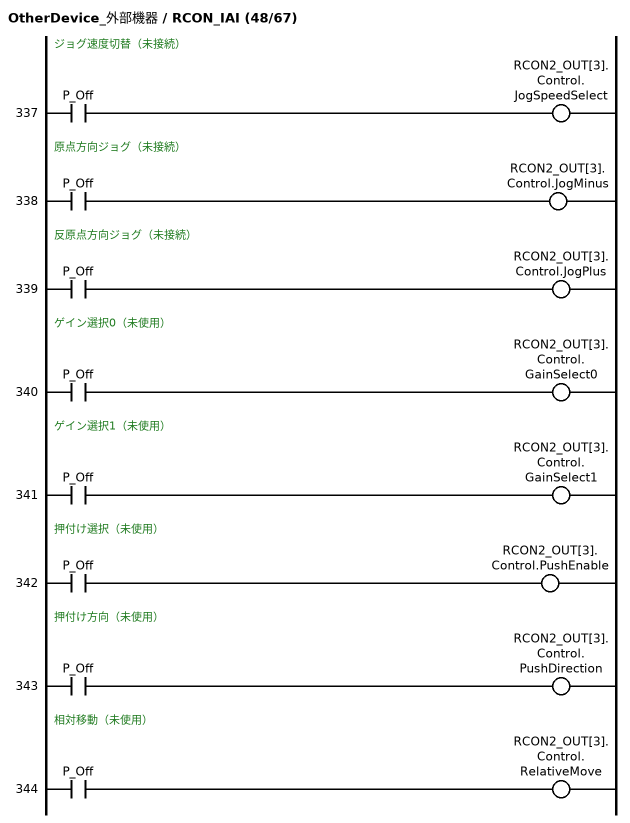
(* Rung 337: ジョグ速度切替（未接続） *)
RCON2_OUT[3].Control.JogSpeedSelect := P_Off;
(* Rung 338: 原点方向ジョグ（未接続） *)
RCON2_OUT[3].Control.JogMinus := P_Off;
(* Rung 339: 反原点方向ジョグ（未接続） *)
RCON2_OUT[3].Control.JogPlus := P_Off;
(* Rung 340: ゲイン選択0（未使用） *)
RCON2_OUT[3].Control.GainSelect0 := P_Off;
(* Rung 341: ゲイン選択1（未使用） *)
RCON2_OUT[3].Control.GainSelect1 := P_Off;
(* Rung 342: 押付け選択（未使用） *)
RCON2_OUT[3].Control.PushEnable := P_Off;
(* Rung 343: 押付け方向（未使用） *)
RCON2_OUT[3].Control.PushDirection := P_Off;
(* Rung 344: 相対移動（未使用） *)
RCON2_OUT[3].Control.RelativeMove := P_Off;

